// SIMATIC S7-200 project (STEP 7-Micro/WIN), CPU 226 CN REL 02.01

SYMBOL_TABLE USUARIO1
ANTI_HORARIO     Q0.4     // Giro del brazo en sentido antihorario
HORARIO          Q0.5     // Giro del brazo en sentido horario
CIL_DOBLE        Q0.6     // Extencion del brazo neumatico
ELEVACION        Q0.3     // Elevacion del brazo neumatico
PINZA_ABIERTA    Q1.0     // Pinza abierta del brazo neumatico
PINZA_CERRADA    Q0.7     // Pinza cerrada del brazo neumatico
DIRECCION_MOTOR  Q0.1     // Drceccion del motor (adelante o atras)
HL1              Q1.5     // Lampara de señalizacion amarilla
HL2              Q1.6     // Lampara de señaliacion verde
HL3              Q1.7     // Lampara de señalizacion roja
CIL_ABAJO        I0.3     // Sensor indicador de cilindro abajo
CIL_ARRIBA       I0.4     // Sensor indicador de cilindro arriba
CIL_EXT          I0.7     // Sensor indicador de cilindro doble extendido
CIL_RET          I1.0     // Sensor indicador de cilindro doble retraido
PINZA_CERRADO    I1.1     // Sensor indicador de Pinza cerrada
ROT_DER          I0.6     // Sensor indicador de cilindro rotatorio a la derecha
ROT_IZQ          I0.5     // Sensor indicador de cilindro rotatorio a la izquierda
FIN_CARRERA_IZQ  I0.2     // Final de carrera izquierda
FIN_CARRERA_DER  I0.1     // Final de carrera derecha
INDUCTIVO        I0.0     // Sensor inductivo
E0               M0.0     // Estado 0
E0a              M1.4     // Estado 0a
E1               M0.1     // Estado 1
E2               M0.2     // Estado 2
E3               M0.3     // Estado 3
E4               M0.4     // Estado 4
E5               M0.5     // Estaro 5
E6               M0.6     // Estado 6
E7               M0.7     // Estado 7
E8               M1.0     // Estado 8
E9               M1.1     // Estado 9
S1               M1.2     // Estado S1
S2               M1.3     // Estado S2
SBB1             I2.5     // Pulsador de marcha
SBB2             I2.4     // Pulsador de paro
SA               I2.7     // Selector rotativo
QS               I2.6     // Zeta de emergencia
FIN_MOV_1        V50.0    // Posicion de memoria para almacenar el movimiento lineal del brazo neumatico 1
FIN_MOV_2        V50.1    // Posicion de memoria para almacenar el movimiento lineal del brazo neumatico 2
FIN_MOV_3        V50.2    // Posicion de memoria para almacenar el movimiento lineal del brazo neumatico 3
FIN_MOV_4        V50.3    // Posicion de memoria para almacenar el movimiento lineal del brazo neumatico 4
FIN_MOV_5        V50.4    // Posicion de memoria para almacenar el movimiento lineal del brazo neumatico 5
FIN_MOV_6        V50.5    // Posicion de memoria para almacenar el movimiento lineal del brazo neumatico 6
FIN_MOV_7        V50.6    // Posicion de memoria para almacenar el movimiento lineal del brazo neumatico 7
EA               M1.5     // Estado EA
M1               M1.6     // Estado M1
M2               M1.7     // Estado M2
M3               M2.0     // Estado M3
M4               M2.1     // Estado M4
M5               M2.2     // Estado M5
SAA              M2.3     // Estado SAA
EB               M2.4     // Estado EB
M6               M2.5     // Estado M6
M7               M2.6     // Estado M7
M8               M2.7     // Estado M8
M9               M3.0     // Estado M9
M10              M3.1     // Estado M10
M11              M3.2     // Estado M11
M12              M3.3     // Estado M12
M13              M3.4     // Estado M13
M14              M3.5     // Estado M14
M15              M3.6     // Estado M15
M16              M3.7     // Estado M16
M17              M4.0     // Estado M17
SB               M4.1     // Estado SB
EC               M4.2     // Estado EC
M18              M4.3     // Estado M18
M19              M4.4     // Estado M19
M20              M4.5     // Estado M20
M21              M4.6     // Estado M21
M22              M4.7     // Estado M22
M23              M5.0     // Estado M23
M24              M5.1     // Estado M24
M25              M5.2     // Estado M25
M26              M5.3     // Estado M26
M27              M5.4     // Estado M27
M28              M5.5     // Estado M28
M29              M5.6     // Estado M29
SC               M5.7     // Estado SC
E_D              M6.0     // Estado E_D
M30              M6.1     // Estado M30
M31              M6.2     // Estado M31
M32              M6.3     // Estado M32
M33              M6.4     // Estado M33
SD               M6.5     // Estado SD
ciclo            M7.0     // Bit de indicacion para la comunicacion
error_comunica   M7.1     // Bit indicador si hay error en la comunicacion
GO_ALIMENTACION  V0.0     // Iniciar la unidad de alimentacion desde la unidad de transporte
GO_ENSAMBLAJE    V0.2     // Iniciar la unidad de ensamblaje desde la unidad de transporte
GO_PROCESAMIENTO V0.4     // Iniciar la unidad de procesamiento desde la unidad de transporte
GO_SELECCION     V0.6     // Iniciar la unidad de seleccion desde la unidad de transporte
FIN_ALIMENTACION V1.1     // Indica la finalizacion de la unidad y asi el brazo recoja los cilindros
FIN_ENSAMBLAJE   V2.3     // Indica la finalizacion de la unidad y asi el brazo recoja los cilindros
FIN_PROCESAMIENTO V3.5     // Indica la finalizacion de la unidad y asi el brazo recoja los cilindros
EE1              M7.2     // Estado EE1
EE2              M7.3     // Estado EE2
EE3              M7.4     // Estado EE3
MMA              M7.5     // Estado MMA
EEE              M7.6     // Estado EEE
END_SYMBOL_TABLE

ORGANIZATION_BLOCK PRINCIPAL:OB1
TITLE=COMENTARIOS DEL PROGRAMA
BEGIN
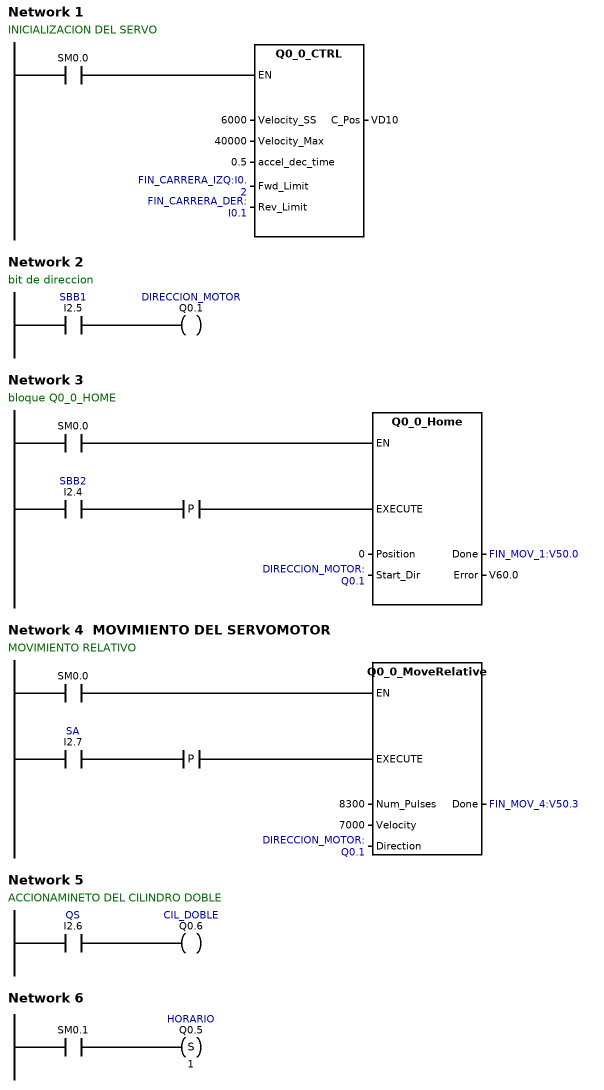
Network 1
// INICIALIZACION DEL SERVO
LD     SM0.0
CALL   Q0_0_CTRL:SBR1, 6000, 40000, 0.5, FIN_CARRERA_IZQ:I0.2, FIN_CARRERA_DER:I0.1, VD10
Network 2
// bit de direccion
LD     SBB1:I2.5
=      DIRECCION_MOTOR:Q0.1
Network 3
// bloque Q0_0_HOME
// (network saved uncompiled; LAD cells follow)
// row 0: c0 -| |- SM0.0  c1 --  c2 --  c3 [Q0_0_Home EN:=power@row0, EXECUTE:=power@row1, Position:=0, Start_Dir:=DIRECCION_MOTOR:Q0.1, Done=>FIN_MOV_1:V50.0, Error=>V60.0]
// row 1: c0 -| |- SBB2:I2.4  c1 -|P|-  c2 --  c3 [box]
// row 2: c3 [box]
Network 4 // MOVIMIENTO DEL SERVOMOTOR
// MOVIMIENTO RELATIVO
LD     SM0.0
=      L60.0
LD     SA:I2.7
EU
=      L63.7
LD     L60.0
CALL   Q0_0_MoveRelative:SBR4, L63.7, 8300, 7000, DIRECCION_MOTOR:Q0.1, FIN_MOV_4:V50.3
Network 5
// ACCIONAMINETO DEL CILINDRO DOBLE
LD     QS:I2.6
=      CIL_DOBLE:Q0.6
Network 6
LD     SM0.1
S      HORARIO:Q0.5, 1
END_ORGANIZATION_BLOCK

// SBR1: protected block, not included

// SBR2: protected block, not included

// SBR3: protected block, not included

// SBR4: protected block, not included

// SBR5: protected block, not included

// SBR6: protected block, not included

// SBR7: protected block, not included

// SBR11: protected block, not included
